(* IEC 61131-3 sources: helmsman/crates/helmsman-canvas/src/fixtures/pump-station, 7 files *)

(* ---- analog_scale.st ---- *)
(* Raw analog count to engineering units, held to the range. bad is set when
   the raw value is outside raw_min..raw_max by more than the margin: a broken
   wire on a 4-20 mA loop, or a transmitter that has failed. *)
FUNCTION_BLOCK analog_scale
VAR_INPUT
  raw : REAL;
  raw_min : REAL := 0.0;
  raw_max : REAL := 32767.0;
  eng_min : REAL := 0.0;
  eng_max : REAL := 100.0;
  margin : REAL := 0.05;
END_VAR
VAR_OUTPUT
  value : REAL;
  bad : BOOL;
END_VAR
VAR
  span : REAL;
END_VAR
span := raw_max - raw_min;
bad := span <= 0.0 OR raw < raw_min - span * margin OR raw > raw_max + span * margin;
IF span > 0.0 THEN
  value := LIMIT(eng_min, eng_min + (raw - raw_min) / span * (eng_max - eng_min), eng_max);
END_IF;
END_FUNCTION_BLOCK

(* ---- duty_standby.st ---- *)
(* Two machines sharing one job. The duty unit runs on demand; the standby
   runs when asked to assist or when the duty unit is not available. Duty
   swaps at every stop, so both wear evenly. *)
FUNCTION_BLOCK duty_standby
VAR_INPUT
  demand : BOOL;
  assist : BOOL;
  a_ok : BOOL;
  b_ok : BOOL;
END_VAR
VAR_OUTPUT
  run_a : BOOL;
  run_b : BOOL;
  b_is_duty : BOOL;
  none_available : BOOL;
END_VAR
VAR
  stopped : F_TRIG;
END_VAR
stopped(CLK := demand);
IF stopped.Q THEN
  b_is_duty := NOT b_is_duty;
END_IF;
IF b_is_duty THEN
  run_b := demand AND b_ok;
  run_a := demand AND a_ok AND (assist OR NOT b_ok);
ELSE
  run_a := demand AND a_ok;
  run_b := demand AND b_ok AND (assist OR NOT a_ok);
END_IF;
none_available := demand AND NOT a_ok AND NOT b_ok;
END_FUNCTION_BLOCK

(* ---- latched_alarm.st ---- *)
(* One alarm: on after on_delay, stays showing until the condition has gone
   and someone has acknowledged it. *)
FUNCTION_BLOCK latched_alarm
VAR_INPUT
  condition : BOOL;
  ack : BOOL;
  on_delay : TIME;
END_VAR
VAR_OUTPUT
  active : BOOL;
  unacked : BOOL;
  showing : BOOL;
END_VAR
VAR
  delay : TON;
  rise : R_TRIG;
END_VAR
delay(IN := condition, PT := on_delay);
active := delay.Q;
rise(CLK := active);
IF rise.Q THEN
  unacked := TRUE;
ELSIF ack THEN
  unacked := FALSE;
END_IF;
showing := active OR unacked;
END_FUNCTION_BLOCK

(* ---- main.st ---- *)
(* Lift station: two pumps on one wet well, duty and standby, run from a level
   transmitter between start and stop levels. The standby assists at a higher
   level and takes over from a pump that has faulted; duty swaps at each stop.

   plant_model.st stands in for the well and pumps so this runs with nothing
   wired. To wire real I/O: delete plant_model.st, delete the plant lines in
   the PROGRAM (each one says PLANT), and point io.map at your remote I/O
   module.

   A hardwired high-level float and motor protection belong in hardware;
   nothing here is a safety function. *)

(* Turns the well level into demand, assist and the level alarms. *)
FUNCTION_BLOCK well_control
VAR_INPUT
  level_m : REAL;
  level_bad : BOOL;
  low_float : BOOL;
  ack : BOOL;
END_VAR
VAR_OUTPUT
  demand : BOOL;
  assist : BOOL;
  dry_run_lockout : BOOL;
  alarm_new : BOOL;
  alarm_showing : BOOL;
END_VAR
VAR CONSTANT
  stop_at_m : REAL := 0.8;
  start_at_m : REAL := 2.0;
  assist_at_m : REAL := 2.6;
  high_at_m : REAL := 3.4;
  dry_at_m : REAL := 0.3;
END_VAR
VAR
  high : latched_alarm;
  dry : latched_alarm;
  transmitter : latched_alarm;
END_VAR
IF level_m >= start_at_m THEN
  demand := TRUE;
ELSIF level_m <= stop_at_m THEN
  demand := FALSE;
END_IF;
IF level_m >= assist_at_m THEN
  assist := TRUE;
ELSIF level_m <= start_at_m THEN
  assist := FALSE;
END_IF;
high(condition := level_m >= high_at_m, ack := ack, on_delay := T#5s);
dry(condition := low_float OR level_m <= dry_at_m, ack := ack, on_delay := T#0s);
transmitter(condition := level_bad, ack := ack, on_delay := T#2s);
dry_run_lockout := dry.active OR transmitter.active;
alarm_new := high.unacked OR dry.unacked OR transmitter.unacked;
alarm_showing := high.showing OR dry.showing OR transmitter.showing;
END_FUNCTION_BLOCK

FUNCTION_BLOCK pump_pair
VAR_INPUT
  demand : BOOL;
  assist : BOOL;
  ack : BOOL;
  fb_a : BOOL;
  fb_b : BOOL;
  overload_a : BOOL;
  overload_b : BOOL;
END_VAR
VAR_OUTPUT
  contactor_a : BOOL;
  contactor_b : BOOL;
  alarm_new : BOOL;
  alarm_showing : BOOL;
END_VAR
VAR
  duty : duty_standby;
  pump_a : motor_starter;
  pump_b : motor_starter;
  pump_fault : latched_alarm;
  none_left : latched_alarm;
END_VAR
duty(demand := demand, assist := assist, a_ok := NOT pump_a.fault, b_ok := NOT pump_b.fault);
pump_a(run := duty.run_a, feedback := fb_a, overload := overload_a, reset := ack);
pump_b(run := duty.run_b, feedback := fb_b, overload := overload_b, reset := ack);
pump_fault(condition := pump_a.fault OR pump_b.fault, ack := ack, on_delay := T#0s);
none_left(condition := duty.none_available, ack := ack, on_delay := T#0s);
contactor_a := pump_a.contactor;
contactor_b := pump_b.contactor;
alarm_new := pump_fault.unacked OR none_left.unacked;
alarm_showing := pump_fault.showing OR none_left.showing;
END_FUNCTION_BLOCK

PROGRAM pump_station
VAR_INPUT
  start_pb : BOOL;
  stop_pb : BOOL;
  ack_pb : BOOL;
  fb_a_in : BOOL;
  fb_b_in : BOOL;
  overload_a_in : BOOL;
  overload_b_in : BOOL;
  low_float_in : BOOL;
END_VAR
VAR_OUTPUT
  pump_a : BOOL;
  pump_b : BOOL;
  lamp_green : BOOL;
  lamp_red : BOOL;
  level_m : REAL;
END_VAR
VAR
  plant : plant_model;  (* PLANT *)
  level_tx : analog_scale;
  well : well_control;
  pumps : pump_pair;
  light : stack_light;
  run : BOOL;
  level_raw : REAL;
  fb_a : BOOL;
  fb_b : BOOL;
END_VAR

plant(pump_a := pump_a, pump_b := pump_b);  (* PLANT *)
level_raw := plant.level_raw;  (* PLANT: read your analog input here *)
fb_a := fb_a_in OR plant.fb_a;  (* PLANT: keep the _in input *)
fb_b := fb_b_in OR plant.fb_b;  (* PLANT: keep the _in input *)
run := (run OR start_pb) AND NOT stop_pb;

level_tx(raw := level_raw, eng_min := 0.0, eng_max := 4.0);
well(level_m := level_tx.value, level_bad := level_tx.bad, low_float := low_float_in, ack := ack_pb);
pumps(demand := run AND well.demand AND NOT well.dry_run_lockout,
      assist := well.assist, ack := ack_pb, fb_a := fb_a, fb_b := fb_b,
      overload_a := overload_a_in, overload_b := overload_b_in);
light(running := run, alarm_new := well.alarm_new OR pumps.alarm_new,
      alarm_showing := well.alarm_showing OR pumps.alarm_showing);

pump_a := pumps.contactor_a;
pump_b := pumps.contactor_b;
lamp_green := light.green;
lamp_red := light.red;
level_m := level_tx.value;
END_PROGRAM

(* ---- motor_starter.st ---- *)
(* Motor starter with contactor feedback and a latched fault.
   feedback is the contactor's auxiliary contact, overload the thermal relay.
   fault_code: 0 none, 1 overload, 2 no feedback after a start or feedback
   lost while running, 3 feedback with no command (contactor stuck on).
   A fault drops the contactor and holds until reset. An emergency stop
   belongs in a hardwired safety circuit, not in this block. *)
FUNCTION_BLOCK motor_starter
VAR_INPUT
  run : BOOL;
  feedback : BOOL;
  overload : BOOL;
  reset : BOOL;
  feedback_time : TIME := T#2s;
END_VAR
VAR_OUTPUT
  contactor : BOOL;
  running : BOOL;
  fault : BOOL;
  fault_code : INT;
END_VAR
VAR
  no_feedback : TON;
  stuck_on : TON;
END_VAR
no_feedback(IN := contactor AND NOT feedback, PT := feedback_time);
stuck_on(IN := NOT contactor AND feedback, PT := feedback_time);
IF overload THEN
  fault_code := 1;
ELSIF no_feedback.Q THEN
  fault_code := 2;
ELSIF stuck_on.Q THEN
  fault_code := 3;
ELSIF reset THEN
  fault_code := 0;
END_IF;
fault := fault_code <> 0;
contactor := run AND NOT fault;
running := contactor AND feedback;
END_FUNCTION_BLOCK

(* ---- plant_model.st ---- *)
(* PLANT MODEL: not part of the controls. Stands in for the wet well and the
   pumps so the program moves with nothing wired. Inflow alternates between
   dry and storm weather. Delete this file when you wire real I/O. *)
FUNCTION_BLOCK plant_model
VAR_INPUT
  pump_a : BOOL;
  pump_b : BOOL;
END_VAR
VAR_OUTPUT
  level_raw : REAL;
  fb_a : BOOL;
  fb_b : BOOL;
END_VAR
VAR CONSTANT
  dry_inflow : REAL := 0.01;      (* m/s of well level *)
  storm_inflow : REAL := 0.06;
  pump_outflow : REAL := 0.03;    (* m/s of well level, each pump *)
  weather_change : TIME := T#2m;
  motor_delay : TIME := T#500ms;
  dt_s : REAL := 0.1;
END_VAR
VAR
  motor_a : TON;
  motor_b : TON;
  clock : TON;
  weather : TON;
  storm : BOOL;
  level_m : REAL := 1.5;  {state unit=m}
  inflow : REAL;
END_VAR
motor_a(IN := pump_a, PT := motor_delay);
motor_b(IN := pump_b, PT := motor_delay);
fb_a := motor_a.Q;
fb_b := motor_b.Q;

weather(IN := NOT weather.Q, PT := weather_change);
IF weather.Q THEN
  storm := NOT storm;
END_IF;
IF storm THEN
  inflow := storm_inflow;
ELSE
  inflow := dry_inflow;
END_IF;
clock(IN := NOT clock.Q, PT := T#100ms);
IF clock.Q THEN
  level_m := level_m + inflow * dt_s;
  IF fb_a THEN
    level_m := level_m - pump_outflow * dt_s;
  END_IF;
  IF fb_b THEN
    level_m := level_m - pump_outflow * dt_s;
  END_IF;
  level_m := LIMIT(0.0, level_m, 4.0);
END_IF;
level_raw := level_m / 4.0 * 32767.0;
END_FUNCTION_BLOCK

(* ---- stack_light.st ---- *)
(* Green while running. Red flashes for an alarm nobody has acknowledged and
   is steady for one that is acknowledged but still there. *)
FUNCTION_BLOCK stack_light
VAR_INPUT
  running : BOOL;
  alarm_new : BOOL;
  alarm_showing : BOOL;
END_VAR
VAR_OUTPUT
  green : BOOL;
  red : BOOL;
END_VAR
VAR
  flash : BLINK_PATTERN;
  pattern : INT;
END_VAR
IF alarm_new THEN
  pattern := 2;
ELSIF alarm_showing THEN
  pattern := 1;
ELSE
  pattern := 0;
END_IF;
flash(EN := TRUE, MODE := pattern, PERIOD := T#1s);
green := running;
red := flash.Q;
END_FUNCTION_BLOCK
